// TIA Portal V21 export
// export: Created 2026-11-21T13:00:31.875841Z, ExportSetting WithDefaults, DisplayName Totally Integrated Automation Portal, DisplayVersion V21, DisplayName STEP 7 Professional, DisplayVersion V21, DisplayName STEP 7 Safety, DisplayVersion V21, DisplayName Tech WebApplication, DisplayVersion V21, DisplayName WinCC Basic/Comfort/Advanced, DisplayVersion V21, DisplayName WinCC Unified, DisplayVersion V21
PlcWatchTable "Tank"
  PlcWatchTableEntry ""Start""  DisplayFormat=Bool, ModifyTrigger=Permanent, MonitorTrigger=Permanent
  PlcWatchTableEntry ""Setpoint""  DisplayFormat=DEC_signed, ModifyTrigger=Permanent, ModifyValue=50, MonitorTrigger=Permanent, Comment="Half full"
  PlcWatchTableEntry ""Speed""  DisplayFormat=Float, ModifyTrigger=Permanent, ModifyValue=1.5, MonitorTrigger=Permanent
  PlcWatchTableEntry ""StatusWord""  DisplayFormat=Hex, ModifyTrigger=Permanent, MonitorTrigger=OnceOnlyAtStart
  PlcTableCommentEntry   Comment="The recipe"
  PlcWatchTableEntry ""Recipe".count"  DisplayFormat=DEC_signed, ModifyTrigger=Permanent, MonitorTrigger=Permanent
  PlcWatchTableEntry ""Recipe".limits.high"  DisplayFormat=DEC_signed, ModifyTrigger=OnceOnlyAtStart, ModifyValue=85, MonitorTrigger=Permanent
  PlcWatchTableEntry ""Recipe".steps[1].target"  DisplayFormat=Float, ModifyTrigger=Permanent, MonitorTrigger=Permanent
  PlcWatchTableEntry   Address=%MW40, DisplayFormat=Bin, ModifyTrigger=Permanent, MonitorTrigger=Permanent, Comment="No tag at this address"
  PlcWatchTableEntry ""LadBoxesData".sum"  DisplayFormat=DEC_signed, ModifyTrigger=Permanent, MonitorTrigger=Permanent
